// TIA Portal V20 export
// export: Created 2026-10-12T15:48:33.6641892Z, ExportSetting WithDefaults, DisplayName Totally Integrated Automation Portal, DisplayVersion V20, DisplayName TIA Portal Openness, DisplayVersion V20, DisplayName TIA Portal Teamcenter Gateway, DisplayVersion V20, DisplayName TIA Portal Version Control Interface, DisplayVersion V20, DisplayName SINAMICS Startdrive Advanced, DisplayVersion V20 SP1 Update 2, DisplayName SINAMICS Startdrive G110M, G120, G120C, G120D, G120P, G115D, DisplayVersion V20 SP1 Update 2, DisplayName SINAMICS Startdrive G130, G150, S120, S150, SINAMICS MV, G220, S200, S210, DisplayVersion V20 SP1 Update 2, DisplayName STEP 7 Professional, DisplayVersion V20, DisplayName STEP 7 Safety, DisplayVersion V20, DisplayName WinCC Basic/Comfort/Advanced, DisplayVersion V20, DisplayName WinCC Professional, DisplayVersion V20, DisplayName WinCC Unified, DisplayVersion V20
FUNCTION "FRK_ConfigStatus" : Void   // FC108, SCL
{ S7_Optimized_Access := 'TRUE' }
VERSION : 0.1
// stored: AutoNumber true, IsIECCheckEnabled false, SetENOAutomatically false, UDAEnableTagReadback false
   VAR_INPUT
      RootIndex : Int;
      Scope : String;
      PolicyLost : Bool;
      UsersLost : Bool;
   END_VAR
   VAR_IN_OUT
      Persist : "ST_ConfigPersistStatus";
      AlarmLog : "FRK_AlarmLog";
   END_VAR
   VAR_TEMP
      Diag : "ST_Diagnostic";
      Accepted : Bool;
   END_VAR
BEGIN

   IF #RootIndex < 1 OR #RootIndex > 2 THEN
       RETURN;
   END_IF;
   #Persist.Pending := FALSE;
   #Persist.Failed := "FRK_ConfigRuntime".Failed[#RootIndex];
   #Persist.StoreKind := 0;
   // Named set operations are not wired by the live retained-value provider.
   #Persist.StorePresent := TRUE;
   #Persist.RestoreLost := "FRK_ConfigStore".Lost[#RootIndex] OR #PolicyLost OR #UsersLost;
   #Persist.RestoreAcknowledged := "FRK_ConfigStore".Acknowledged[#RootIndex] AND NOT #PolicyLost AND NOT #UsersLost;
   IF #PolicyLost THEN
       #Persist.LostPath := CONCAT(IN1 := #Scope, IN2 := '.AccessPolicy');
   ELSIF #UsersLost THEN
       #Persist.LostPath := CONCAT(IN1 := #Scope, IN2 := '.Access');
   ELSE
       #Persist.LostPath := "FRK_ConfigStore".LostPath[#RootIndex];
   END_IF;
   // Access owns its precise loss events; announce only typed-config loss here.
   IF "FRK_ConfigStore".Lost[#RootIndex] AND NOT "FRK_ConfigStore".Acknowledged[#RootIndex] THEN
       IF "FRK_ConfigRuntime".LossSlot[#RootIndex] = 0 THEN
           #Diag := "FRK_UnitScratch".EmptyDiagnostic;
           #Diag.ReasonCode := 2040;
           #Diag.Description := WSTRING#'std.error.configRestoreLost';
           #Diag.SourcePath := STRING_TO_WSTRING("FRK_ConfigStore".LostPath[#RootIndex]);
           "FRK_ConfigRuntime".LossSlot[#RootIndex] := "FRK_AlarmRaise"(AlarmLog := #AlarmLog, Diag := #Diag, ResetClass := 0);
       END_IF;
   ELSIF "FRK_ConfigRuntime".LossSlot[#RootIndex] > 0 THEN
       #Accepted := "FRK_AlarmGone"(AlarmLog := #AlarmLog, Slot := "FRK_ConfigRuntime".LossSlot[#RootIndex]);
       "FRK_ConfigRuntime".LossSlot[#RootIndex] := 0;
   END_IF;
END_FUNCTION
